// TIA Portal V20 export
Screen "Robot_NBG_Kuka"  1276x673
  ScreenItem "Zone01" at 662,80 size 482x510  Type=HmiGraphicView
  ScreenItem "permanentareaborderrectangle" at 0,0 size 0x0  Type=HmiRectangle
  ScreenItem "Line_Header_X0_Y64" at 0,64 size 1276x0  Type=HmiLine
  ScreenItem "nbgMessages" at 10,479 size 428x169  Type=HmiAlarmControl
  ScreenItem "Robot Name" at 390,3 size 500x37  Type=HmiIOField
  ScreenItem "Button_Back" at 2,2 size 90x60  Type=HmiButton
  ScreenItem "Select NBG" at 390,3 size 500x37  Type=HmiSymbolicIOField
  ScreenItem "Rectangle TG1 Status" at 196,0 size 217x132  Type=HmiRectangle
  ScreenItem "Text field TG1 Status" at 196,0 size 218x31  Type=HmiTextBox
  ScreenItem "Rectangle NBG Status" at 0,0 size 196x178  Type=HmiRectangle
  ScreenItem "Text Field Motor On" at 5,81 size 90x21  Type=HmiTextBox
  ScreenItem "Text Field On Path" at 5,127 size 90x21  Type=HmiTextBox
  ScreenItem "Text Filed E- Stop" at 99,35 size 90x21  Type=HmiTextBox
  ScreenItem "Text Field System Fault" at 99,58 size 90x21  Type=HmiTextBox
  ScreenItem "Text Field Move Pause" at 99,104 size 90x21  Type=HmiTextBox
  ScreenItem "Text Field In Cycle" at 5,104 size 90x21  Type=HmiTextBox
  ScreenItem "Text Field Ready" at 5,58 size 90x21  Type=HmiTextBox
  ScreenItem "Text Field Fault" at 99,81 size 90x21  Type=HmiTextBox
  ScreenItem "Text Field Auto Mode" at 5,35 size 90x21  Type=HmiTextBox
  ScreenItem "Text Field Enable Motion" at 5,150 size 90x21  Type=HmiTextBox
  ScreenItem "Text field NBG Status" at 0,0 size 196x31  Type=HmiTextBox
  ScreenItem "Text Field Full Speed_2" at 99,127 size 90x21  Type=HmiTextBox
  ScreenItem "Text Field TG1 Moving" at 202,35 size 100x21  Type=HmiTextBox
  ScreenItem "Text Field TG1 Move Pause" at 202,58 size 100x21  Type=HmiTextBox
  ScreenItem "Text Field TG1 Fault" at 202,81 size 100x21  Type=HmiTextBox
  ScreenItem "Text Field TG1 With Fixture" at 202,104 size 100x21  Type=HmiTextBox
  ScreenItem "Text Field TG1 ATI Connection" at 306,35 size 100x21  Type=HmiTextBox
  ScreenItem "Text Field TG1 ATI Deconnection" at 306,58 size 100x21  Type=HmiTextBox
  ScreenItem "Text Field TG1 Lock Pos" at 306,81 size 100x21  Type=HmiTextBox
  ScreenItem "Text Field TG1 Unlock Pos" at 306,104 size 100x21  Type=HmiTextBox
  ScreenItem "Rectangle TGA" at 0,0 size 102x91  Type=HmiRectangle
  ScreenItem "Text Field TGA Moving" at 5,3 size 90x21  Type=HmiTextBox
  ScreenItem "Text Field TGA Move Pause" at 5,23 size 90x21  Type=HmiTextBox
  ScreenItem "Text Field TGA Fault" at 5,43 size 90x21  Type=HmiTextBox
  ScreenItem "Text field TGA Status" at 28,68 size 44x21  Type=HmiTextBox
  ScreenItem "Rectangle TGAA" at 102,0 size 282x91  Type=HmiRectangle
  ScreenItem "Text Field TGAA In Storage Pos" at 198,3 size 90x21  Type=HmiTextBox
  ScreenItem "Text Field TGAA In Delivery Pos" at 287,3 size 90x21  Type=HmiTextBox
  ScreenItem "Text Field TGAA With Fixture" at 109,3 size 90x21  Type=HmiTextBox
  ScreenItem "Text field TGAA Status" at 104,68 size 47x21  Type=HmiTextBox
  ScreenItem "Rectangle TGAA Delivery Pos" at 290,29 size 85x56  Type=HmiRectangle
  ScreenItem "Button TGAA Go Delivery Pos" at 291,30 size 83x54  Type=HmiButton
  ScreenItem "TGAA Delivery Pos Interlock" at 0,0 size 100x30  Type=HmiCircle
  ScreenItem "Rectangle TGAA Storage Pos" at 157,29 size 85x56  Type=HmiRectangle
  ScreenItem "Button TGAA Go Storage Pos" at 158,30 size 83x54  Type=HmiButton
  ScreenItem "TGAA Storage Pos Interlock" at 0,0 size 100x30  Type=HmiCircle
  ScreenItem "Rectangle TGB" at 0,0 size 102x91  Type=HmiRectangle
  ScreenItem "Text Field TGB Moving" at 6,3 size 90x21  Type=HmiTextBox
  ScreenItem "Text Field TGB Move Pause" at 6,23 size 90x21  Type=HmiTextBox
  ScreenItem "Text Field TGB Fault" at 6,43 size 90x21  Type=HmiTextBox
  ScreenItem "Text field TGB Status" at 29,68 size 44x21  Type=HmiTextBox
  ScreenItem "Rectangle TGBA" at 102,0 size 282x91  Type=HmiRectangle
  ScreenItem "Text Field TGBA In Storage Pos" at 198,3 size 90x21  Type=HmiTextBox
  ScreenItem "Text Field TGBA In Delivery Pos" at 287,3 size 90x21  Type=HmiTextBox
  ScreenItem "Text Field TGBA With Fixture" at 109,3 size 90x21  Type=HmiTextBox
  ScreenItem "Text field TGBA Status" at 104,68 size 47x21  Type=HmiTextBox
  ScreenItem "Rectangle TGBA Storage Pos" at 157,29 size 85x56  Type=HmiRectangle
  ScreenItem "Rectangle TGBA Delivery Pos" at 290,29 size 85x56  Type=HmiRectangle
  ScreenItem "Button TGBA Go Storage Pos" at 158,30 size 83x54  Type=HmiButton
  ScreenItem "TGBA Storage Pos Interlock" at 0,0 size 100x30  Type=HmiCircle
  ScreenItem "Button TGBA Go Delivery Pos" at 291,30 size 83x54  Type=HmiButton
  ScreenItem "TGBA Delivery Pos Interlock" at 0,0 size 100x30  Type=HmiCircle
  ScreenItem "Rectangle TGAB" at 0,0 size 281x91  Type=HmiRectangle
  ScreenItem "Text Field TGAB In Storage Pos" at 95,3 size 90x21  Type=HmiTextBox
  ScreenItem "Text Field TGAB In Delivery Pos" at 6,3 size 90x21  Type=HmiTextBox
  ScreenItem "Text Field TGAB With Fixture" at 184,3 size 90x21  Type=HmiTextBox
  ScreenItem "Text field TGAB Status" at 233,68 size 47x21  Type=HmiTextBox
  ScreenItem "Rectangle TGAB Delivery Pos" at 9,29 size 85x56  Type=HmiRectangle
  ScreenItem "Button TGAB Go Delivery Pos" at 10,30 size 83x54  Type=HmiButton
  ScreenItem "TGAB Delivery Pos Interlock" at 0,0 size 100x30  Type=HmiCircle
  ScreenItem "Rectangle TGAB Storage Pos" at 142,29 size 85x56  Type=HmiRectangle
  ScreenItem "Button TGAB Go Storage Pos" at 143,30 size 83x54  Type=HmiButton
  ScreenItem "TGAB Storage Pos Interlock" at 0,0 size 100x30  Type=HmiCircle
  ScreenItem "Rectangle TGBB" at 0,0 size 281x91  Type=HmiRectangle
  ScreenItem "Text Field TGBB In Storage Pos" at 95,3 size 90x21  Type=HmiTextBox
  ScreenItem "Text Field TGBB In Delivery Pos" at 6,3 size 90x21  Type=HmiTextBox
  ScreenItem "Text Field TGBB With Fixture" at 184,3 size 90x21  Type=HmiTextBox
  ScreenItem "Text field TGBB Status" at 233,68 size 47x21  Type=HmiTextBox
  ScreenItem "Rectangle TGBB Storage Pos" at 142,29 size 85x56  Type=HmiRectangle
  ScreenItem "Rectangle TGBB Delivery Pos" at 9,29 size 85x56  Type=HmiRectangle
  ScreenItem "Button TGBB Go Storage Pos" at 143,30 size 83x54  Type=HmiButton
  ScreenItem "TGBB Storage Pos Interlock" at 0,0 size 100x30  Type=HmiCircle
  ScreenItem "Button TGBB Go Delivery Pos" at 10,30 size 83x54  Type=HmiButton
  ScreenItem "TGBB Delivery Pos Interlock" at 0,0 size 100x30  Type=HmiCircle
  ScreenItem "Rectangle TGCB" at 0,0 size 281x91  Type=HmiRectangle
  ScreenItem "Text Field TGCB In Storage Pos" at 95,3 size 90x21  Type=HmiTextBox
  ScreenItem "Text Field TGCB In Delivery Pos" at 6,3 size 90x21  Type=HmiTextBox
  ScreenItem "Text Field TGCB With Fixture" at 184,3 size 90x21  Type=HmiTextBox
  ScreenItem "Text field TGCB Status" at 233,68 size 47x21  Type=HmiTextBox
  ScreenItem "Rectangle TGCB Storage Pos" at 142,29 size 85x56  Type=HmiRectangle
  ScreenItem "Rectangle TGCB Delivery Pos" at 9,29 size 85x56  Type=HmiRectangle
  ScreenItem "Button TGCB Go Storage Pos" at 143,30 size 83x54  Type=HmiButton
  ScreenItem "TGCB Storage Pos Interlock" at 0,0 size 100x30  Type=HmiCircle
  ScreenItem "Button TGCB Go Delivery Pos" at 10,30 size 83x54  Type=HmiButton
  ScreenItem "TGCB Delivery Pos Interlock" at 0,0 size 100x30  Type=HmiCircle
  ScreenItem "Text Field TG1 In Load Pos1" at 0,0 size 90x21  Type=HmiTextBox
  ScreenItem "Rectangle Load Pos1" at 2,25 size 85x56  Type=HmiRectangle
  ScreenItem "Button Go Load Pos1" at 3,26 size 83x54  Type=HmiButton
  ScreenItem "TG1 Load Pos1 Interlock" at 0,0 size 100x30  Type=HmiCircle
  ScreenItem "Text Field TG1 In Storage Pos1" at 0,0 size 90x21  Type=HmiTextBox
  ScreenItem "Rectangle Storage Pos1" at 2,26 size 85x56  Type=HmiRectangle
  ScreenItem "Button Go Storage Pos1" at 3,27 size 83x54  Type=HmiButton
  ScreenItem "TG1 Storage Pos1 Interlock" at 0,0 size 100x30  Type=HmiCircle
  ScreenItem "Text Field TG1 In Storage Pos2" at 0,0 size 90x21  Type=HmiTextBox
  ScreenItem "Rectangle Storage Pos2" at 2,26 size 85x56  Type=HmiRectangle
  ScreenItem "Button Go Storage Pos2" at 3,27 size 83x54  Type=HmiButton
  ScreenItem "TG1 Storage Pos2 Interlock" at 0,0 size 100x30  Type=HmiCircle
  ScreenItem "Text Field TG1 In Storage Pos3" at 0,0 size 90x21  Type=HmiTextBox
  ScreenItem "Rectangle Storage Pos3" at 2,26 size 85x56  Type=HmiRectangle
  ScreenItem "Button Go Storage Pos3" at 3,27 size 83x54  Type=HmiButton
  ScreenItem "TG1 Storage Pos3 Interlock" at 0,0 size 100x30  Type=HmiCircle
  ScreenItem "Rectangle TG1_2" at 0,0 size 281x187  Type=HmiRectangle
  ScreenItem "Text Field TG1 In Work Pos1" at 6,4 size 90x21  Type=HmiTextBox
  ScreenItem "Text Field TG1 In Work Pos2" at 96,4 size 90x21  Type=HmiTextBox
  ScreenItem "Text Field TG1 In Work Pos3" at 186,4 size 90x21  Type=HmiTextBox
  ScreenItem "Text Field TG1 In Work Pos4" at 5,99 size 90x21  Type=HmiTextBox
  ScreenItem "Text Field TG1 In Work Pos5" at 95,99 size 90x21  Type=HmiTextBox
  ScreenItem "Text Field TG1 In Work Pos6" at 187,99 size 90x21  Type=HmiTextBox
  ScreenItem "Rectangle Work Pos2" at 98,29 size 85x56  Type=HmiRectangle
  ScreenItem "Button Go Work Pos2" at 99,30 size 83x54  Type=HmiButton
  ScreenItem "TG1 Work Pos2 Interlock" at 0,0 size 100x30  Type=HmiCircle
  ScreenItem "Rectangle Work Pos3" at 188,29 size 85x56  Type=HmiRectangle
  ScreenItem "Button Go Work Pos3" at 189,30 size 83x54  Type=HmiButton
  ScreenItem "TG1 Work Pos3 Interlock" at 0,0 size 100x30  Type=HmiCircle
  ScreenItem "Rectangle Work Pos4" at 7,124 size 85x56  Type=HmiRectangle
  ScreenItem "Button Go Work Pos4" at 8,125 size 83x54  Type=HmiButton
  ScreenItem "TG1 Work Pos4 Interlock" at 0,0 size 100x30  Type=HmiCircle
  ScreenItem "Rectangle Work Pos5" at 97,124 size 85x56  Type=HmiRectangle
  ScreenItem "Button Go Work Pos5" at 98,125 size 83x54  Type=HmiButton
  ScreenItem "TG1 Work Pos5 Interlock" at 0,0 size 100x30  Type=HmiCircle
  ScreenItem "Rectangle Work Pos6" at 187,124 size 85x56  Type=HmiRectangle
  ScreenItem "Button Go Work Pos6" at 188,125 size 83x54  Type=HmiButton
  ScreenItem "TG1 Work Pos6 Interlock" at 0,0 size 100x30  Type=HmiCircle
  ScreenItem "Rectangle Work Pos1" at 8,29 size 85x56  Type=HmiRectangle
  ScreenItem "Button Go Work Pos1" at 9,30 size 83x54  Type=HmiButton
  ScreenItem "TG1 Work Pos1 Interlock" at 0,0 size 100x30  Type=HmiCircle
  ScreenItem "Rectangle TGC" at 0,0 size 102x91  Type=HmiRectangle
  ScreenItem "Text Field TGC Moving" at 6,3 size 90x21  Type=HmiTextBox
  ScreenItem "Text Field TGC Move Pause" at 6,23 size 90x21  Type=HmiTextBox
  ScreenItem "Text Field TGC Fault" at 6,43 size 90x21  Type=HmiTextBox
  ScreenItem "Text field TGC Status" at 29,68 size 44x21  Type=HmiTextBox
  ScreenItem "Rectangle TGCA" at 102,0 size 282x91  Type=HmiRectangle
  ScreenItem "Text Field TGCA In Storage Pos" at 198,3 size 90x21  Type=HmiTextBox
  ScreenItem "Text Field TGCA In Delivery Pos" at 287,3 size 90x21  Type=HmiTextBox
  ScreenItem "Text Field TGCA With Fixture" at 109,3 size 90x21  Type=HmiTextBox
  ScreenItem "Text field TGCA Status" at 104,68 size 47x21  Type=HmiTextBox
  ScreenItem "Rectangle TGCA Storage Pos" at 157,29 size 85x56  Type=HmiRectangle
  ScreenItem "Rectangle TGCA Delivery Pos" at 290,29 size 85x56  Type=HmiRectangle
  ScreenItem "Button TGCA Go Storage Pos" at 158,30 size 83x54  Type=HmiButton
  ScreenItem "TGCA Storage Pos Interlock" at 0,0 size 100x30  Type=HmiCircle
  ScreenItem "Button TGCA Go Delivery Pos" at 291,30 size 83x54  Type=HmiButton
  ScreenItem "TGCA Delivery Pos Interlock" at 0,0 size 100x30  Type=HmiCircle
